FUNCTION_BLOCK SKILL_Condition_BOOL (* One comparison in a decision of a skill (for example Weight greater than 1.9): answers YES or NO. Technical: Compares Operand with Expected by Operator (eq, ne): YES or NO *)
  (* Standard: 61499-2 *)
  (* Version 0.1, 2026-09-28, Project contributors, AAU Smart Production Lab *)
  PACKAGE modlib;
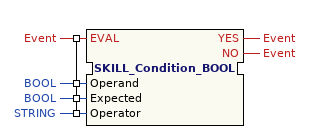
  EVENT_INPUT
    EVAL WITH Operand, Expected, Operator; (* Evaluate the condition (the steps before it are done) *)
  END_EVENT
  EVENT_OUTPUT
    YES; (* The condition holds: the first branch *)
    NO; (* The condition does not hold: the second branch, or past the conditional steps *)
  END_EVENT
  VAR_INPUT
    Operand : BOOL; (* What is compared: a parameter of the skill or a result of a step *)
    Expected : BOOL; (* What it is compared with *)
    Operator : STRING := 'eq'; (* eq, ne, gt, gte, lt or lte: Operand <op> Expected *)
  END_VAR
  VAR
    Holds : BOOL;
  END_VAR
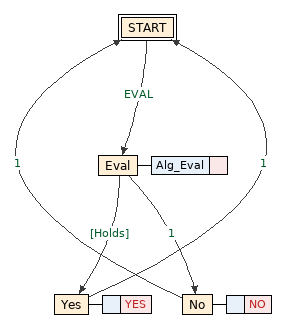
  EC_STATES
    START;
    Eval : Alg_Eval;
    Yes : -> YES;
    No : -> NO;
  END_STATES
  EC_TRANSITIONS
    START TO Eval := EVAL;
    Eval TO Yes := [Holds];
    Eval TO No := 1;
    Yes TO START := 1;
    No TO START := 1;
  END_TRANSITIONS
  ALGORITHM Alg_Eval IN ST:
Holds := ((Operator = 'eq') AND (Operand = Expected)) OR ((Operator = 'ne') AND (Operand <> Expected));
  END_ALGORITHM
END_FUNCTION_BLOCK
